//静止状态 road相同,分road分方向讨论
IF (_pPremover^.stAxisStatus.nNcCycleCounter=0)THEN      //premover is not ready
    IF 	(_pPremover^.stNcTOPLC.nCuRoadID=stRoad1_Param.nRoadID)THEN
		 IF (_eDirection=E_Direction.DIRECTION_POSITIVE)THEN
			_fPrePosition:=_pPremover^.stNcTOPLC.fActPos-_pPremover^.stAxisParam.fClampLength*0.5-_fGap;
			IF _bIsGroupMember THEN   //03.31
				_fPrePosition:=_pPremover^.stNcTOPLC.fActPos-_fGroupInGap;
				IF _pPremover^.stPLCTONC.bEndPosCalDone AND(stAxis.stAxisStatus.nNcCycleCounter=0)THEN   //04.03
					_fPrePosition:=_pPremover^.stPLCTONC.stEndPosition.fPosition-_fGroupInGap;
				END_IF
			END_IF
		 ELSE
			_fPrePosition:=_pPremover^.stNcTOPLC.fActPos+_pPremover^.stAxisParam.fClampLength*0.5+_fGap;
			IF _bIsGroupMember THEN   //03.31
				_fPrePosition:=_pPremover^.stNcTOPLC.fActPos+_fGroupInGap;
				IF _pPremover^.stPLCTONC.bEndPosCalDone AND(stAxis.stAxisStatus.nNcCycleCounter=0)THEN   //04.03
					_fPrePosition:=_pPremover^.stPLCTONC.stEndPosition.fPosition+_fGroupInGap;
				END_IF
			END_IF
		 END_IF
	ELSE
		IF (_eNextRoadDirection=E_Direction.DIRECTION_POSITIVE)THEN
			_fPrePosition:=_pPremover^.stNcTOPLC.fActPos-_pPremover^.stAxisParam.fClampLength*0.5-_fGap;
			IF _bIsGroupMember THEN   //03.31
				_fPrePosition:=_pPremover^.stNcTOPLC.fActPos-_fGroupInGap;
				IF _pPremover^.stPLCTONC.bEndPosCalDone AND(stAxis.stAxisStatus.nNcCycleCounter=0)THEN   //04.03
					_fPrePositionTemp:=_pPremover^.stPLCTONC.stEndPosition.fPosition-_fGroupInGap;
					IF (_fPrePositionTemp>=stRoad2_Param.fEndPosition)THEN
						_fPrePosition:=stRoad2_Param.fEndPosition;
					ELSE
						_fPrePosition:=_pPremover^.stPLCTONC.stEndPosition.fPosition-_fGroupInGap;
					END_IF
				END_IF
			END_IF
		ELSE
			_fPrePosition:=_pPremover^.stNcTOPLC.fActPos+_pPremover^.stAxisParam.fClampLength*0.5+_fGap;
			IF _bIsGroupMember THEN   //03.31
				_fPrePosition:=_pPremover^.stNcTOPLC.fActPos+_fGroupInGap;
				IF _pPremover^.stPLCTONC.bEndPosCalDone AND(stAxis.stAxisStatus.nNcCycleCounter=0)THEN   //04.03
					_fPrePositionTemp:=_pPremover^.stPLCTONC.stEndPosition.fPosition+_fGroupInGap;
					IF (_fPrePositionTemp<=stRoad2_Param.fEndPosition)THEN
						_fPrePosition:=stRoad2_Param.fEndPosition;
					ELSE
						_fPrePosition:=_pPremover^.stPLCTONC.stEndPosition.fPosition+_fGroupInGap;
					END_IF
				END_IF
			END_IF
		END_IF
	END_IF 
	//_bRunning:=FALSE;
END_IF

IF (stAxis.stNcTOPLC.nCuRoadID=stRoad1_Param.nRoadID)THEN    //road1
		IF (_eDirection=E_Direction.DIRECTION_POSITIVE)THEN
			IF (_fPrePosition<=stAxis.stNcTOPLC.fActPos)THEN
			    _bSegOver:=TRUE;
			     RETURN; 
			END_IF
		ELSE
			IF (_fPrePosition>=stAxis.stNcTOPLC.fActPos)THEN
					_bSegOver:=TRUE;
					RETURN; 
			END_IF
		END_IF
		_fNewPrePosition:=_fPrePosition;
		stAxis.stPLCTONC.stEndPosition.nRoadID:=stRoad1_Param.nRoadID; 
ELSE    //road2
		IF (_eNextRoadDirection=E_Direction.DIRECTION_POSITIVE)THEN
			IF (_fPrePosition<=stAxis.stNcTOPLC.fActPos)THEN
					_bSegOver:=TRUE;
					RETURN; 
		    END_IF
		
			IF _fPrePosition>stRoad2_Param.fEndPosition THEN
				_fNewPrePosition:=stRoad2_Param.fEndPosition;
			ELSE
				_fNewPrePosition:=_fPrePosition;
			END_IF
		    
		ELSE
			IF (_fPrePosition>=stAxis.stNcTOPLC.fActPos)THEN
				_bSegOver:=TRUE;
				RETURN; 
			END_IF
			IF _fPrePosition<stRoad2_Param.fEndPosition THEN
				_fNewPrePosition:=stRoad2_Param.fEndPosition;
			ELSE
				_fNewPrePosition:=_fPrePosition;
			END_IF
		END_IF
		stAxis.stPLCTONC.stEndPosition.nRoadID:=stRoad2_Param.nRoadID;
END_IF
_bSegOver:=FALSE;
END_ACTION

ACTION A_StopPathGerenation:

_fPostion:=0.5*stAxis.stNcTOPLC.fActVelo*stAxis.stNcTOPLC.fActVelo/_fDec;

IF stAxis.stAxisStatus.bPositiveDirection THEN
		 IF (stAxis.stNcTOPLC.nCuRoadID=stAxis.stPLCTONC.nRoadID_1) THEN
			 _fStopPosition:=_fPostion+stAxis.stNcTOPLC.fActPos-stAxis.stPLCTONC.fRoad1_Length;
			 IF (_fStopPosition>0) THEN 
				  _fNewStopPosition:=FC_TransformPosition(fOffset:=stAxis.stPLCTONC.fRoad1_Length , fPosition:=_fStopPosition );    //坐标转换
				  stAxis.stPLCTONC.stEndPosition.fPosition:=_fNewStopPosition;
				  
				  stAxis.stPLCTONC.stStartPosition.nRoadID:=stAxis.stPLCTONC.nRoadID_1;
				  stAxis.stPLCTONC.stEndPosition.nRoadID:=stAxis.stPLCTONC.nRoadID_2;
				  
			 ELSE
				 stAxis.stPLCTONC.stEndPosition.fPosition:=_fPostion+stAxis.stNcTOPLC.fActPos;
				 stAxis.stPLCTONC.stStartPosition.nRoadID:=stAxis.stPLCTONC.nRoadID_1;
				 stAxis.stPLCTONC.stEndPosition.nRoadID:=stAxis.stPLCTONC.nRoadID_1;

			 END_IF
		 ELSE
			 
				 IF NOT stAxis.stPLCTONC.bRoadDirection THEN   //04.08
				     stAxis.stPLCTONC.stEndPosition.fPosition:=_fPostion+stAxis.stNcTOPLC.fActPos;
					 IF (stAxis.stPLCTONC.stEndPosition.fPosition>=stAxis.stPLCTONC.fRoad2_Length)THEN
					    _bStopPosError:=TRUE;
				     END_IF 
				 ELSE
					 stAxis.stPLCTONC.stEndPosition.fPosition:=stAxis.stNcTOPLC.fActPos-_fPostion;
					 IF (stAxis.stPLCTONC.stEndPosition.fPosition<=0)THEN
					    _bStopPosError:=TRUE;
				     END_IF
				 END_IF
				 stAxis.stPLCTONC.stStartPosition.nRoadID:=stAxis.stPLCTONC.nRoadID_2;
				 stAxis.stPLCTONC.stEndPosition.nRoadID:=stAxis.stPLCTONC.nRoadID_2;
				 (*IF (stAxis.stPLCTONC.stEndPosition.fPosition>=stAxis.stPLCTONC.fRoad2_Length)OR (stAxis.stPLCTONC.stEndPosition.fPosition<=0)THEN
					 _bStopPosError:=TRUE;
				 END_IF*) 
			 
		 END_IF
ELSE
		IF (stAxis.stNcTOPLC.nCuRoadID=stAxis.stPLCTONC.nRoadID_1) THEN
			 _fStopPosition:=stAxis.stNcTOPLC.fActPos-_fPostion;
			 IF (_fStopPosition<0) THEN 
				  _fNewStopPosition:=FC_TransformPosition(fOffset:=0 , fPosition:=_fStopPosition );    //坐标转换
				  stAxis.stPLCTONC.stEndPosition.fPosition:=_fNewStopPosition;
				  stAxis.stPLCTONC.stStartPosition.nRoadID:=stAxis.stPLCTONC.nRoadID_1;
				  stAxis.stPLCTONC.stEndPosition.nRoadID:=stAxis.stPLCTONC.nRoadID_2;
				 // stAxis.stPLCTONC.nRoadOrder:=0;
			 ELSE
				 stAxis.stPLCTONC.stEndPosition.fPosition:=stAxis.stNcTOPLC.fActPos-_fPostion;
				stAxis.stPLCTONC.stStartPosition.nRoadID:=stAxis.stPLCTONC.nRoadID_1;
				 stAxis.stPLCTONC.stEndPosition.nRoadID:=stAxis.stPLCTONC.nRoadID_1;
			 END_IF
		 ELSE
			 (*stAxis.stPLCTONC.stEndPosition.fPosition:=stAxis.stNcTOPLC.fActPos-_fPostion;
	         stAxis.stPLCTONC.stStartPosition.nRoadID:=stAxis.stPLCTONC.nRoadID_2;
			 stAxis.stPLCTONC.stEndPosition.nRoadID:=stAxis.stPLCTONC.nRoadID_2;
			 IF (stAxis.stPLCTONC.stEndPosition.fPosition<=0)THEN
				 _bStopPosError:=TRUE;
			 END_IF *)
			 IF NOT stAxis.stPLCTONC.bRoadDirection THEN   //04.08
				     stAxis.stPLCTONC.stEndPosition.fPosition:=_fPostion+stAxis.stNcTOPLC.fActPos;
					 IF (stAxis.stPLCTONC.stEndPosition.fPosition>=stAxis.stPLCTONC.fRoad2_Length)THEN
					    _bStopPosError:=TRUE;
				     END_IF 
			 ELSE
					 stAxis.stPLCTONC.stEndPosition.fPosition:=stAxis.stNcTOPLC.fActPos-_fPostion;
					 IF (stAxis.stPLCTONC.stEndPosition.fPosition<=0)THEN
					    _bStopPosError:=TRUE;
				     END_IF
		     END_IF
			 stAxis.stPLCTONC.stStartPosition.nRoadID:=stAxis.stPLCTONC.nRoadID_2;
			 stAxis.stPLCTONC.stEndPosition.nRoadID:=stAxis.stPLCTONC.nRoadID_2;
			 
		 END_IF
END_IF


stAxis.stPLCTONC.fTargetVelocity:=stAxis.stNcTOPLC.fActVelo;
stAxis.stPLCTONC.stEndPosition.fVelocity:=0;
stAxis.stPLCTONC.stEndPosition.fAccleration:=_fDec;
stAxis.stPLCTONC.stEndPosition.fDeceleration:=_fDec;
END_ACTION

ACTION A_UpstateStatus:
stAxis.stAxisStatus.nCycleCounter:=_nCycleCount;
stAxis.stAxisStatus.bCollisionStoped:=_bCollisionChecked;
//02.24
_nLastCycleCounter:=_nCycleCount;
_nLastNcCycleCounter:=stAxis.stAxisStatus.nNcCycleCounter_WP;

IF (_nStep=0)THEN 
	RETURN;
END_IF

(*IF (stAxis.stNcTOPLC.nCuRoadID<>stRoad1_Param.nRoadID)AND NOT _bAddNodeOk  THEN 
	IF stAxis.stPLCTONC.bRoadDirection THEN   //负向头部
		_bAddNodeOk:=_fbAxisGroupList.M_AddNode(aRoadRef:=GVL_MC.aRoadRef , bHeadNode:=TRUE , nRoadId:=stRoad2_Param.nRoadID , pAixs:=ADR(stAxis));
	ELSE
		_bAddNodeOk:=_fbAxisGroupList.M_AddNode(aRoadRef:=GVL_MC.aRoadRef , bHeadNode:=FALSE , nRoadId:=stRoad2_Param.nRoadID , pAixs:=ADR(stAxis));
	END_IF
 
END_IF
IF (stAxis.stNcTOPLC.nCuRoadID<>stRoad1_Param.nRoadID)AND  NOT _bDeleteNodeOk THEN 
  
   _bDeleteNodeOk:=_fbAxisGroupList.M_DeleteNode(aRoadRef:=GVL_MC.aRoadRef , nSysType:=stAxis.stPLCTONC.nSysType , nRoadId:=stRoad1_Param.nRoadID , pAixs:=ADR(stAxis) );
     
END_IF*)  //04.14注释
// 04.14修改 防止fork更新前置后 后置更新错误
(*IF (_stRoad1_Param.nRoadID<>0)THEN
	IF (stAxis.stNcTOPLC.nCuRoadID<>_stRoad1_Param.nRoadID)AND NOT _bAddNodeOk  THEN 
		IF stAxis.stPLCTONC.bRoadDirection THEN   //负向头部
			_bAddNodeOk:=_fbAxisGroupList.M_AddNode(aRoadRef:=GVL_MC.aRoadRef , bHeadNode:=TRUE , nRoadId:=stRoad2_Param.nRoadID , pAixs:=ADR(stAxis));
		ELSE
			_bAddNodeOk:=_fbAxisGroupList.M_AddNode(aRoadRef:=GVL_MC.aRoadRef , bHeadNode:=FALSE , nRoadId:=stRoad2_Param.nRoadID , pAixs:=ADR(stAxis));
		END_IF
	 
	END_IF
	IF (stAxis.stNcTOPLC.nCuRoadID<>_stRoad1_Param.nRoadID)AND  NOT _bDeleteNodeOk THEN 
	  
	   _bDeleteNodeOk:=_fbAxisGroupList.M_DeleteNode(aRoadRef:=GVL_MC.aRoadRef , nSysType:=stAxis.stPLCTONC.nSysType , nRoadId:=stRoad1_Param.nRoadID , pAixs:=ADR(stAxis) );
		 
	END_IF
END_IF*)
END_ACTION

END_FUNCTION_BLOCK

(* stored: Version 1.1.0.1, ProductVersion 3.1.4024.12
   POU FTS_MCMoveAbsoluteForkCA: Id {bb3928c7-0f5b-43c3-94fd-7501df7a2b60}, SpecialFunc None
   Action A_CommandCheck: Id {95859b2c-f943-4273-9a2c-f0f4275a5af5}
   Action A_DyPathDisCal: Id {5521bf29-cc71-406a-88db-ab2a0f2fab53}
   Action A_DyPathDisCalTans: Id {d16b9390-ebeb-4505-b358-71799a4a6bb8}
   Action A_DyPathDisCalTansLast: Id {20a22e23-acc9-4224-a1a0-eaeec7d6b572}
   Action A_DyPathDisCalTansPre: Id {0dce8342-54c5-4c45-8944-3cb8926e2732}
   Action A_Init: Id {3237e363-c5de-41cd-b1a9-dd8d32dd1181}
   Action A_MeasureIn: Id {f264282a-0798-4f5d-93b8-e5c3924a5de8}
   Action A_NextMoverCheck: Id {d71a99b2-61a9-4f43-942f-886a5b66b97c}
   Action A_NextPathMoverUpdateCheck: Id {3f0f7f34-d1d7-41de-ae9f-7fd48a41c92c}
   Action A_NextPathUpdateCheck: Id {e10756a5-6ae5-449e-92a3-c1dcdbf74a79}
   Action A_ParamCheck: Id {a14eeaef-ea2d-42e8-a36e-5d28e828bd13}
   Action A_PathPreGeneration: Id {f91c7592-121a-456e-81fe-90300b19219b}
   Action A_PathUpdateCheck: Id {ff4afa3d-2d83-4102-8672-76e170cc92e7}
   Action A_PreMoverCheck: Id {77e8e3d0-4818-419f-a086-2b7b54c356bd}
   Action A_PreMoverCheckForkCmd: Id {07ebacf6-6a9a-4770-a98e-16fae82ebab5}
   Action A_PreMoverCheckNotForkCmd: Id {e779d5df-f3d0-4018-8f15-b1a3ec2790ca}
   Action A_StopPathGerenation: Id {40ef551d-e417-46d3-86da-8c71edf95abc}
   Action A_UpstateStatus: Id {ff0037ef-e6b4-4015-8807-f9a63e00864b} *)
